SUBAPPLICATION Remote_Init_Retry (* INIT fuer einen Remote-OPC-UA-Client: INITO sofort an die Kette, bei INITO- neuer Versuch nach DT *)
  (* Standard: 61499-2; Description: Copyright (c) 2026 Meisterschulen am Ostbahnhof This program and the accompanying materials are made available under the terms of the Eclipse Public License 2.0 which is available at https://www.eclipse.org/legal/epl-2.0/ SPDX-License-Identifier: EPL-2.0 *)
  (* Version 1.1, 2026-10-30, Franz Höpfinger, Meisterschulen am Ostbahnhof, INIT-FB (events::init::INIT) direkt hinter dem Eingang INIT: SubApp wird im fboot aufgeloest, ohne ihn bliebe bei unverbundenem INIT nur E_MERGE_2.EI1 (Event, kein EInit) und E_TRIG loeste nie aus. Jetzt bleibt ein EInit-Eingang, unverbunden wird er automatisch ausgeloest. *)
  (* Version 1.0, 2026-10-30, Franz Höpfinger, Meisterschulen am Ostbahnhof, Neu. forte (#1092): Remote-Client meldet INITO+ erst wenn der Node existiert, sonst nach Timeout INITO- und Stopp, neuer Versuch nur durch neues INIT+. Abgestimmt mit ELFMASTER: E_DELAY vor erneutem INIT+, bei INIT mit QI=FALSE E_DELAY.STOP, reagiert auf jedes INITO-. *)
  PACKAGE MyLib::sys;
  (* Documentation:
  Neuer Versuch fuer einen Remote-OPC-UA-Client
   Seit forte #1092 meldet ein Remote-Client (SUBSCRIBE/WRITE/CALL_METHOD auf eine andere Station) INITO+ erst, wenn der Node auf der Gegenstation existiert. Sonst kommt nach dem Timeout (Standard 60 s) INITO- und der Client versucht es nicht mehr von selbst.
    - INIT geht sofort an den Client (CLIENT_INIT) und gleich als INITO weiter: die Kette wartet nicht auf die Gegenstation.
   - Kommt vom Client INITO mit QO=FALSE und ist QI=TRUE, wird nach DT (Standard 2 s) erneut INIT gesendet - bei jedem INITO-, nicht nur beim ersten.
   - INIT mit QI=FALSE stoppt eine laufende Pause.
   - INIT darf unverbunden bleiben: der innere events::init::INIT haelt im fboot einen EInit-Eingang, E_TRIG loest ihn aus.
    Verdrahtung: CLIENT_INIT an Client.INIT, Client.INITO an CLIENT_INITO, Client.QO an CLIENT_QO, QI gemeinsam. Nur fuer Remote-Clients einsetzen, nicht in den Adapter-Huellen selbst.
  *)
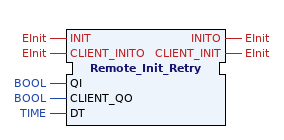
  EVENT_INPUT
    INIT : EInit; (* INIT aus der Kette (QI wie am Client) *)
    CLIENT_INITO : EInit; (* INITO des Remote-Clients *)
  END_EVENT
  EVENT_OUTPUT
    INITO : EInit; (* Sofort nach INIT, wartet nicht auf den Client *)
    CLIENT_INIT : EInit; (* An INIT des Remote-Clients *)
  END_EVENT
  VAR_INPUT
    QI : BOOL := TRUE; (* Gleiches QI wie am Client *)
    CLIENT_QO : BOOL; (* QO des Remote-Clients *)
    DT : TIME := T#2s; (* Pause vor neuem Versuch *)
  END_VAR
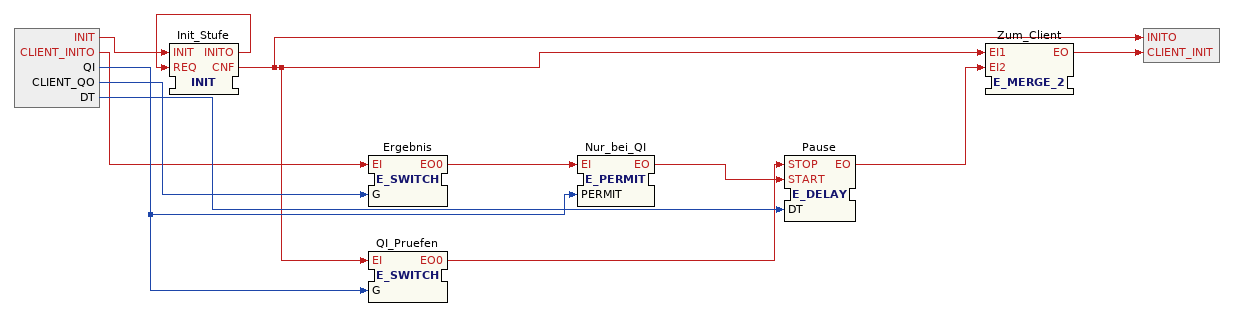
  FBS
    Init_Stufe : events::init::INIT; (* Haelt den EInit-Eingang im fboot (E_TRIG) *)
    QI_Pruefen : iec61499::events::E_SWITCH; (* INIT mit QI=FALSE stoppt eine laufende Pause *)
    Ergebnis : iec61499::events::E_SWITCH; (* EO0: INITO- (QO=FALSE) *)
    Nur_bei_QI : iec61499::events::E_PERMIT;
    Pause : iec61499::events::E_DELAY;
    Zum_Client : iec61499::events::E_MERGE_2; (* erster Versuch + Neuversuche *)
  END_FBS
  EVENT_CONNECTIONS
    INIT TO Init_Stufe.INIT;
    Init_Stufe.INITO TO Init_Stufe.REQ;
    Init_Stufe.CNF TO Zum_Client.EI1;
    Init_Stufe.CNF TO INITO;
    Init_Stufe.CNF TO QI_Pruefen.EI;
    QI_Pruefen.EO0 TO Pause.STOP;
    CLIENT_INITO TO Ergebnis.EI;
    Ergebnis.EO0 TO Nur_bei_QI.EI;
    Nur_bei_QI.EO TO Pause.START;
    Pause.EO TO Zum_Client.EI2;
    Zum_Client.EO TO CLIENT_INIT;
  END_CONNECTIONS
  DATA_CONNECTIONS
    QI TO QI_Pruefen.G;
    CLIENT_QO TO Ergebnis.G;
    QI TO Nur_bei_QI.PERMIT;
    DT TO Pause.DT;
  END_CONNECTIONS
END_SUBAPPLICATION
